Staubli VAL3: bind.pgx

public program bind()
  local string l_sbtn
  local num l_i
begin
  userPageBindClick("point","btnback",bBack,true)
  userPageBind("point","lbl2","innerHTML",sTrajItem,1,"r")
  userPageBind("point","lbllib","innerHTML",sUsingLib,1,"r")
  userPageBind("point","lblframe","innerHTML",sUsingFrame,1,"r")
  userPageBind("point","lbltool","innerHTML",sUsingTool,1,"r")

  userPageBind("point","lblpageindex","innerHTML",sPageIndex,1,"r")
  userPageBind("point","lblpagenum","innerHTML",sPageNum,1,"r")

  //click
  for l_i = 0 to size(bBool)-1
    l_sbtn="btn"+toString("",l_i)
    userPageBindClick("point",l_sbtn,bBool[l_i],true)
  endFor

  //lst
  //userPageBind("point","lst1","options",sList,49,"r")

  userPageBind("point","lst1","value",sSelPoint,1,"rw")
end
